Fanuc KAREL source: NC0062.compact.KL

PROGRAM NC0062
%STACKSIZE=65535
%PRIORITY=65535
%NOLOCKGROUP
ROUTINE R FROM NC0062
ROUTINE R
VAR
S1 : INTEGER
S2 : INTEGER
BEGIN
S1=1
FOR S2=1 TO 2 DO
S1=(S1 + 1)
ENDFOR
END R
BEGIN
R
END NC0062
